(* IEC 61131-3 sources: plcassist-cli/packages/volt-lsp-iec/test-corpus/pro2193/Device/Plc Logic/Application/99 Library/Function Blocks/Actuators/Pumps, 3 files *)

(* ---- LubricationPumpFB.fb ---- *)
// ---------- Lubrication pump control ------------
{attribute 'symbol' := 'none'}
FUNCTION_BLOCK LubricationPumpFB
EXTENDS ActuatorWithAlarm_BaseFB
IMPLEMENTS IActuator
VAR_INPUT
	xEnable					: BOOL;		// Enable the lubrication pump (Machine is running in automatic mode)
	{attribute 'symbol' := 'read'}	xPulseInput				: BOOL;		// Input: When the pump is running, count the number of pulses on this input
	errorId					: WORD;
END_VAR
VAR_IN_OUT
	RunningTime				: UDINT;	// Map as persistent var (je mag geen retain vars gebruiken in FB's, daarom als IN_OUT var)
	NumberOfStarts			: UDINT;	// Map as persistent var
	iHoursCounter			: INT;		// Count hours until next lubrication
	iInterval				: INT;		// Start lubricating after this many hours
END_VAR
VAR//VISU
	{attribute 'symbol' := 'readwrite'}	xTestLubrication		: BOOL;		// Manually test the lubrication from the Keba panel
	{attribute 'symbol' := 'read'}		iPulseCounter			: INT;		// Show the number of counted pulses on the panel
	{attribute 'symbol' := 'read'}		xPumpRunning			: BOOL;		// High when vacuum pump output is high
END_VAR
VAR
	Pump					: ActuatorFB;
	NoPulseAlarm			: SetErrorFB;

	T_1Hour					: BTON;
	T_Lubricate				: BTON;
	Trig_StartPump			: TriggerFB;
	Trig_TestLubrication	: TriggerFB;
	Trig_Input				: TriggerFB;
END_VAR
VAR CONSTANT
	rLubricationPumpLength	: REAL := 2 * 60;		// Lubrication pump will run for this time after each interval. Default is 2 minutes.
END_VAR

SUPER^();

xPumpRunning			:= Pump.Map();
iInterval				:= MAX(iInterval, 1);	// Interval must be at least 1 hour.
NoPulseAlarm.alarmCondition	:= FALSE;

IF T_1Hour.Set(xEnable, 60 * 60) THEN	// Gives a trigger output once every hour.
	iHoursCounter		:= iHoursCounter + 1;
	T_1Hour.Reset();
END_IF

IF Trig_StartPump.Rising(iHoursCounter >= iInterval) THEN
	Pump.Set();
	iPulseCounter		:= 0;
END_IF

IF xPumpRunning AND Trig_Input.AnyEdge(xPulseInput) THEN
	Increment.AnyInt(iPulseCounter);
END_IF

IF T_Lubricate.Set(In := xPumpRunning, Pt := rLubricationPumpLength) THEN
	iHoursCounter		:= 0;
	Pump.Reset();
	NoPulseAlarm.alarmCondition := iPulseCounter = 0;
END_IF

IF Trig_TestLubrication.Rising(xTestLubrication) THEN
	IF xPumpRunning THEN
		iHoursCounter	:= 0;
		NoPulseAlarm.alarmCondition := iPulseCounter = 0;
	ELSE
		iPulseCounter	:= 0;
	END_IF
	Pump.SetOrReset(NOT xPumpRunning);
END_IF

NoPulseAlarm(
	moduleHandler	:= moduleHandler,
	textRefId		:= textRefId,
	alarmCondition	:= ,
	alarmDelay		:= alarmDelay,
	errorId			:= errorId,
	severity		:= severity,
	reaction		:= reaction,
	active			=> );

Pump();

// ---------- Measure total running time and number of starts of lubrication pump ------------
//CalcOnTime(
//	xIn			:= xPumpRunning,
//	xReset		:= ,
//	uliSeconds	:= RunningTime,
//	uliCycles	:= NumberOfStarts);

END_FUNCTION_BLOCK

METHOD PROTECTED Alarms
END_METHOD

// Maps the actuator to the physical output
METHOD PUBLIC Map : BOOL
Map := Pump.Map();
END_METHOD

// Reset the output (=False)
METHOD PUBLIC Reset
Pump.Reset();
END_METHOD

{attribute 'hide'}
METHOD PUBLIC Set : BOOL
// no implementation
END_METHOD

{attribute 'hide'}
METHOD PUBLIC SetOrReset
VAR_INPUT
	xValue	: BOOL;
END_VAR
// no implementation
END_METHOD

(* ---- VacuumPumpDualFB.fb ---- *)
// Control a vacuum pump configuration with individual pumps for high and low vacuum
FUNCTION_BLOCK VacuumPumpDualFB
EXTENDS ActuatorWithAlarm_BaseFB
IMPLEMENTS IActuator
VAR_INPUT
	xMachineRunning				: BOOL;		// Machine is running in automatic mode
	xMainAirValve				: BOOL;		// Main air valve is switched on
	xManualOnOffSwitch			: BOOL;
	xThermalInputHighVacuum		: BOOL;		// Input: High when thermal contact switched
	xThermalInputLowVacuum		: BOOL;		// Input: High when thermal contact switched
	xPhaseCheck					: BOOL;		// Input: High when the fases are in order
	xLowVacuumtankFull			: BOOL;		// Input: Low vacuum tank is full
	xHighVacuumtankFull			: BOOL;		// Input: High vacuum tank is full
	xOptionDisableWithAirButton	: BOOL;		// Map as persistent variable. Option to also disable pump together with main air valve.
	xOptionDisableVacuumPumps	: BOOL;		// Map as presistent variable. Option to disable vacuum pump 2 (Low) and run only High vacuum
	xOptionDisableVacuumPump2	: BOOL;		// Map as presistent variable. Option to disable vacuum pump 2 (Low) and run only High vacuum

	errorId_PhaseCheck			: WORD;		// G_dwAlarms.05	0005 - Three-phase power in wrong order. Change phase connection.
	errorId_Thermal				: WORD;		// G_dwAlarms.06	0006 - Thermal contact Vacuum pump switch off.
	errorId_TooMuchRequested	: WORD;		// G_dwAlarms.07	0007 - Too much vacuum requested. Vacuum level dropped.
	errorId_HighTankDoesNotFill	: WORD;		// G_dwAlarms.13	0013 - Takes too long before high vacuum tank is full.
	errorId_Maintenance			: WORD;		// G_dwWarnings.28	0428 - Warnings: Vacuum Pump ≥  3000 hours of operation. Check manual for maintenance.
END_VAR
VAR_IN_OUT
	TotalRunningTime			: UDINT;	// Map as persistent var (je mag geen retain vars gebruiken in FB's, daarom als IN_OUT var)
	TotalNumberOfStarts			: UDINT;	// Map as persistent var
END_VAR
VAR_OUTPUT
	xVacuumpumpRunning			: BOOL;		// High when vacuum pump output is high
END_VAR
VAR
	HighVacuumPump				: VacuumPumpFB;
	LowVacuumPump				: VacuumPumpFB;
	TotalRunningTime2			: UDINT;	// Not used
	TotalNumberOfStarts2		: UDINT;	// Not used
END_VAR

HighVacuumPump(
	moduleHandler				:= moduleHandler,
	textRefId					:= textRefId,
	alarmEnable					:= alarmEnable,
	alarmDelay					:= alarmDelay,
	severity					:= severity,
	reaction					:= reaction,
	xMachineRunning				:= xMachineRunning,
	xMainAirValve				:= xMainAirValve,
	xManualOnOffSwitch			:= xManualOnOffSwitch,
	xThermalInput				:= xThermalInputHighVacuum,
	xPhaseCheck					:= xPhaseCheck,
	xLowVacuumtankFull			:= xLowVacuumtankFull,
	xHighVacuumtankFull			:= xHighVacuumtankFull,
	xOptionDisableWithAirButton	:= xOptionDisableWithAirButton,
	xOptionDisableVacuumPump	:= xOptionDisableVacuumPumps,
	errorId_PhaseCheck			:= errorId_PhaseCheck,
	errorId_Thermal				:= errorId_Thermal,
	errorId_TooMuchRequested	:= errorId_TooMuchRequested,
	errorId_HighTankDoesNotFill	:= errorId_HighTankDoesNotFill,
	errorId_Maintenance			:= errorId_Maintenance,
	TotalRunningTime			:= TotalRunningTime,
	TotalNumberOfStarts			:= TotalNumberOfStarts,
	xVacuumpumpRunning			=> );

LowVacuumPump(
	moduleHandler				:= moduleHandler,
	textRefId					:= textRefId,
	alarmEnable					:= alarmEnable,
	alarmDelay					:= alarmDelay,
	severity					:= severity,
	reaction					:= reaction,
	xMachineRunning				:= xMachineRunning,
	xMainAirValve				:= xMainAirValve,
	xManualOnOffSwitch			:= xManualOnOffSwitch,
	xThermalInput				:= xThermalInputLowVacuum,
	xPhaseCheck					:= xPhaseCheck,
	xLowVacuumtankFull			:= xLowVacuumtankFull,
	xHighVacuumtankFull			:= xHighVacuumtankFull,
	xOptionDisableWithAirButton	:= xOptionDisableWithAirButton,
	xOptionDisableVacuumPump	:= xOptionDisableVacuumPumps OR xOptionDisableVacuumPump2,
	errorId_PhaseCheck			:= errorId_PhaseCheck,
	errorId_Thermal				:= errorId_Thermal,
	errorId_TooMuchRequested	:= errorId_TooMuchRequested,
	errorId_HighTankDoesNotFill	:= errorId_HighTankDoesNotFill,
	errorId_Maintenance			:= errorId_Maintenance,
	TotalRunningTime			:= TotalRunningTime2,
	TotalNumberOfStarts			:= TotalNumberOfStarts2,
	xVacuumpumpRunning			=> );

xVacuumpumpRunning	:= HighVacuumPump.xVacuumpumpRunning
					OR LowVacuumPump.xVacuumpumpRunning
					OR xOptionDisableVacuumPumps;

END_FUNCTION_BLOCK

METHOD PROTECTED Alarms
END_METHOD

// Maps the actuator to the physical output
{attribute 'hide'}
METHOD PUBLIC Map : BOOL
// no implementation
END_METHOD

// Maps the actuator to the physical output
METHOD PUBLIC MapHigh : BOOL
MapHigh := HighVacuumPump.Map();
END_METHOD

// Maps the actuator to the physical output
METHOD PUBLIC MapLow : BOOL
MapLow := LowVacuumPump.Map();
END_METHOD

// Maps the actuator to the physical output
METHOD PUBLIC MapSwitchTanks : BOOL
MapSwitchTanks := LowVacuumPump.MapSwitchTanks();
END_METHOD

// Reset the output (=False)
METHOD PUBLIC Reset
HighVacuumPump.Reset();
LowVacuumPump.Reset();
END_METHOD

{attribute 'hide'}
METHOD PUBLIC Set : BOOL
// no implementation
END_METHOD

{attribute 'hide'}
METHOD PUBLIC SetOrReset
VAR_INPUT
	xValue	: BOOL;
END_VAR
// no implementation
END_METHOD

(* ---- VacuumPumpFB.fb ---- *)
// Control a standard vacuum pump configuration
FUNCTION_BLOCK VacuumPumpFB
EXTENDS ActuatorWithAlarm_BaseFB
IMPLEMENTS IActuator
VAR_INPUT
	xMachineRunning				: BOOL;		// Machine is running in automatic mode
	xMainAirValve				: BOOL;		// Main air valve is switched on
	xManualOnOffSwitch			: BOOL;
	xThermalInput				: BOOL;		// Input: High when thermal contact switched
	xPhaseCheck					: BOOL;		// Input: High when the fases are in correct order
	xLowVacuumtankFull			: BOOL;		// Input: Low vacuum tank is full
	xHighVacuumtankFull			: BOOL;		// Input: High vacuum tank is full
	xOptionDisableWithAirButton	: BOOL;		// Map as persistent variable. Option to also disable pump together with main air valve.
	xOptionDisableVacuumPump	: BOOL;		// Map as presistent variable. Option to disable vacuum pump 2 (Low) and run only High vacuum

	errorId_PhaseCheck			: WORD;		// G_dwAlarms.05	0005 - Three-phase power in wrong order. Change phase connection.
	errorId_Thermal				: WORD;		// G_dwAlarms.06	0006 - Thermal contact Vacuum pump switch off.
	errorId_TooMuchRequested	: WORD;		// G_dwAlarms.07	0007 - Too much vacuum requested. Vacuum level dropped.
	errorId_HighTankDoesNotFill	: WORD;		// G_dwAlarms.13	0013 - Takes too long before high vacuum tank is full.
	errorId_Maintenance			: WORD;		// G_dwWarnings.28	0428 - Warnings: Vacuum Pump ≥  3000 hours of operation. Check manual for maintenance.
END_VAR
VAR_IN_OUT
	TotalRunningTime			: UDINT;	// Map as persistent var (je mag geen retain vars gebruiken in FB's, daarom als IN_OUT var)
	TotalNumberOfStarts			: UDINT;	// Map as persistent var
END_VAR
VAR_OUTPUT
	xVacuumpumpRunning			: BOOL;		// High when vacuum pump output is high
END_VAR
VAR
	VacuumPump					: ActuatorFB;
	SwitchVacuumTanks			: ActuatorFB;
	PhaseCheckAlarm				: SetErrorFB;
	ThermalAlarm				: SetErrorFB;
	TooMuchRequestedAlarm		: SetErrorFB;
	HighTankDoesNotFillAlarm	: SetErrorFB;
	MaintenanceAlarm			: SetErrorFB;

	Trig_OnOffSwitch			: RisingTriggerFB;
	Trig_MainAirValve			: TriggerFB;
	Trig_StartVacuum			: RisingTriggerFB;
	xVacuumReached				: BOOL;
END_VAR
VAR CONSTANT
	udiVacuumPumpServiceInterval: UDINT := 3000;	// Service interval for vacuum pumps. Default is 3000 hours or 1 year, whichever comes first.
END_VAR

SUPER^();

Trig_MainAirValve.Call(xMainAirValve);
VacuumPump();
SwitchVacuumTanks();
xVacuumpumpRunning	:= VacuumPump.Map();

IF PhaseCheckAlarm.active OR ThermalAlarm.active OR xOptionDisableVacuumPump THEN
	VacuumPump.Reset();
ELSE
	IF xOptionDisableWithAirButton THEN
		IF Trig_MainAirValve.Q_Rising THEN	// Vacuumpump goes on at the same time as the main air valve.
			VacuumPump.Set();
		END_IF
		IF Trig_MainAirValve.Q_Falling THEN	// Reset op luchtknop als Functie actief is anders alleen op tijd of noodstop.
			VacuumPump.Reset();
		END_IF
	END_IF
	IF xMachineRunning THEN
		VacuumPump.Set();
	ELSE
		IF Trig_OnOffSwitch.Rising(xManualOnOffSwitch) THEN
			VacuumPump.SetOrReset(NOT xVacuumpumpRunning);
		END_IF
	END_IF
END_IF

// Alarm wordt pas gegenereerd als er minimaal 1 keer hoog vacuum is gezien.
xVacuumReached		S= Trig_StartVacuum.Rising(xVacuumpumpRunning AND xHighVacuumtankFull);
xVacuumReached		R= NOT xVacuumpumpRunning;

// ---------- Measure total running time and number of starts of vacuum pump ------------
VacuumPump.MeasureOnTime.SetExternalSecondsReference(TotalRunningTime);
VacuumPump.MeasureOnTime.SetExternalCyclesReference(TotalNumberOfStarts);

// ---------- Switch pump from low to high vacuum tank (optional) ------------
SwitchVacuumTanks.SetOrReset(xLowVacuumtankFull AND xVacuumpumpRunning);		// When the Low vacuumtank has reached level, switch the pump to the High vacuumtank.

END_FUNCTION_BLOCK

METHOD PROTECTED Alarms
PhaseCheckAlarm(
	moduleHandler	:= moduleHandler,
	textRefId		:= textRefId,
	alarmCondition	:= NOT xPhaseCheck,
	alarmDelay		:= 0.5,
	errorId			:= errorId_PhaseCheck,			// 002 - Change phase.
	severity		:= enumErrorSeverity.Fault,
	reaction		:= enumErrorReaction.FastStop,
	active			=> );

ThermalAlarm(
	moduleHandler	:= moduleHandler,
	textRefId		:= textRefId,
	alarmCondition	:= xThermalInput,
	alarmDelay		:= 1.0,
	errorId			:= errorId_Thermal,				// 007 - Thermal contact Vacuum pump switch off
	severity		:= enumErrorSeverity.Fault,
	reaction		:= enumErrorReaction.EndCycle,
	active			=> );

MaintenanceAlarm(
	moduleHandler	:= moduleHandler,
	textRefId		:= textRefId,
	alarmCondition	:= TotalRunningTime >= udiVacuumPumpServiceInterval * 60 * 60,
	alarmDelay		:= 0.0,
	errorId			:= errorId_Maintenance,			// Maintenance of vacuum pump is required.
	severity		:= enumErrorSeverity.Warning_Lock,
	reaction		:= enumErrorReaction.No_reaction,
	active			=> );

TooMuchRequestedAlarm(
	moduleHandler	:= moduleHandler,
	textRefId		:= textRefId,
	alarmCondition	:= xVacuumReached AND VacuumPump.Map() AND NOT xHighVacuumtankFull,
	alarmDelay		:= alarmDelay,
	errorId			:= errorId_TooMuchRequested,	// Too much vacuum requested. Vacuum level dropped.
	severity		:= severity,
	reaction		:= reaction,
	active			=> );

HighTankDoesNotFillAlarm(
	moduleHandler	:= moduleHandler,
	textRefId		:= textRefId,
	alarmCondition	:= NOT xVacuumReached AND VacuumPump.Map(),
	alarmDelay		:= 60.0,
	errorId			:= errorId_HighTankDoesNotFill,	// 0013 - Takes too long before high vacuum tank is full
	severity		:= severity,
	reaction		:= reaction,
	active			=> );
END_METHOD

// Maps the actuator to the physical output
METHOD PUBLIC Map : BOOL
Map := VacuumPump.Map();
END_METHOD

// Maps the actuator to the physical output
METHOD PUBLIC MapSwitchTanks : BOOL
MapSwitchTanks := SwitchVacuumTanks.Map();
END_METHOD

// Reset the output (=False)
METHOD PUBLIC Reset
VacuumPump.Reset();
END_METHOD

{attribute 'hide'}
METHOD PUBLIC Set : BOOL
// no implementation
END_METHOD

{attribute 'hide'}
METHOD PUBLIC SetOrReset
VAR_INPUT
	xValue	: BOOL;
END_VAR
// no implementation
END_METHOD
